    rq_activate_all_grippers(True)
    # end: URCap Program Node
  end
  $ 55 "zero_ftsensor()"
  zero_ftsensor()
  $ 56 "EXTT"
  $ 57 "Set GRP_3F_Enable=Off"
  set_standard_digital_out(4, False)
  $ 58 "Set BarcodeTrigger=Off"
  set_standard_digital_out(6, False)
  $ 59 "Set GRP_3F_Decap=Off"
  set_standard_digital_out(3, False)
  $ 60 "Set GRP_3F_Cap=Off"
  set_standard_digital_out(2, False)
  $ 61 "Set GRP_3F_Open=Off"
  set_standard_digital_out(5, False)
  $ 62 "PSE_T≔get_tool_free_pose(dir=[0,0,0.150], move_in_base_frame=True)"
  global PSE_T=get_tool_free_pose(dir=[0,0,0.150], move_in_base_frame=True)
  $ 63 "If is_reachable(Base_const, [PSE_T])"
  if (is_reachable(p[0.0,0.0,0.0,0.0,0.0,0.0], [PSE_T])):
    $ 64 "MoveL"
    $ 65 "PSE_T" "breakAfter"
    movel(PSE_T, a=1.2, v=0.15)
  end
  while (True):
    $ 66 "Robot Program"
    $ 67 "MAIN"
    $ 68 "command_manager(external_control='uGO', cond_suspend=(ITM_Manipulated and AMR_AtTarget and AMR_Charging and AMR_Battery<40), cond_unsuspend=(AMR_Battery≟60))"
    command_manager(external_control="uGO", cond_suspend=(ITM_Manipulated  and  AMR_AtTarget  and  AMR_Charging  and  AMR_Battery<40), cond_unsuspend=(AMR_Battery == 60))
    $ 69 "log_state(STATE_Info)"
    log_state(STATE_Info)
    $ 70 "Switch STATE"
    switch_1 = STATE
    $ 71 "Case 1"
    if (1 == switch_1):
      $ 72 "Stopping"
      $ 73 "STATE_Info≔'Stopping'"
      global STATE_Info="Stopping"
      $ 74 "end_freedrive_mode()"
      end_freedrive_mode()
      $ 75 "Set"
      set_tcp(p[0.0,0.0,0.161,3.1415,0.0,0.0])
      $ 76 "PSE_T≔get_tool_free_pose(dir=[0,0,0.150], move_in_base_frame=True)"
      global PSE_T=get_tool_free_pose(dir=[0,0,0.150], move_in_base_frame=True)
      $ 77 "If is_reachable(Base_const, [PSE_T])"
      if (is_reachable(p[0.0,0.0,0.0,0.0,0.0,0.0], [PSE_T])):
        $ 78 "MoveL"
        $ 79 "PSE_T" "breakAfter"
        movel(PSE_T, a=1.2, v=0.15)
      end
      $ 80 "do_transition(keep_rxry=OBJ_Picked, r=0)"
      do_transition(keep_rxry=OBJ_Picked, r=0)
      $ 89 "Call Sub_AMR_MiR_V3"
      Sub_AMR_MiR_V3()
      $ 90 "If stopping() and AMR_Done"
      if (stopping()  and  AMR_Done):
        $ 91 "STATE≔2"
        global STATE=2
        $ 92 "ugo_update_outputs()"
        ugo_update_outputs()
      end
    elif (2 == switch_1):
      $ 93 "Case 2"
      $ 94 "Stopped"
      $ 95 "STATE_Info≔'Stopped'"
      global STATE_Info="Stopped"
      $ 96 "Call Sub_AMR_MiR_V3"
      Sub_AMR_MiR_V3()
      $ 97 "If CMD_Reset"
      if (CMD_Reset):
        $ 98 "STATE≔3"
        global STATE=3
        $ 99 "ugo_update_outputs()"
        ugo_update_outputs()
      end
    elif (3 == switch_1):
      $ 100 "Case 3"
      $ 101 " Resetting"
      $ 102 "STATE_Info≔'Resetting'"
      global STATE_Info="Resetting"
      $ 103 "uML"
      $ 104 "reset_error()"
      reset_error()
      $ 105 "reset_warning()"
      reset_warning()
      $ 106 "PROCESS_Step≔0"
      global PROCESS_Step=0
      $ 107 "PROCESS_Info≔''"
      global PROCESS_Info=""
      $ 108 "ARM_Referenced≔ False "
      global ARM_Referenced=  False
      $ 109 "WRK_Done≔ False "
      global WRK_Done=  False
      $ 110 "ITM_Prepared≔ False "
      global ITM_Prepared=  False
      $ 111 "ITM_Manipulated≔ False "
      global ITM_Manipulated=  False
      $ 112 "STP≔0"
      global STP=0
      $ 113 "Action≔0"
      global Action=0
      $ 114 "Action_Info≔''"
      global Action_Info=""
      $ 115 "ITM_ID≔0"
      global ITM_ID=0
      $ 116 "JIG≔0"
      global JIG=0
      $ 117 "JIG_Slot≔0"
      global JIG_Slot=0
      $ 118 "Task_info≔''"
      global Task_info=""
      $ 119 "Set"
      set_tcp(p[0.0,0.0,0.161,3.1415,0.0,0.0])
      $ 120 "App"
      $ 121 "'ADD APPLICATION SPECIFIC COMMANDS'"
      # 'ADD APPLICATION SPECIFIC COMMANDS'
      $ 122 "OBJ_Type≔0"
      global OBJ_Type=0
      $ 123 "OBJ_Nbr≔0"
      global OBJ_Nbr=0
      $ 124 "If CNT_Rack_Output≥50"
      if (CNT_Rack_Output >= 50):
        $ 125 "CNT_Rack_Output≔0"
        global CNT_Rack_Output=0
      end
      $ 126 "TASK≔struct(ID=0, NAVI=struct(target=0, footprint=0, protectiveOff=0, dock=0), WORK=struct(ITM_ID_Src=0, JIG_ID_Src=0, OBJ_Nbr_Src=0, ACT_Src=0, ITM_ID_Tgt=0, JIG_ID_Tgt=0, OBJ_Nbr_Tgt=0, ACT_Tgt=0, OBJ_Type=0))"
      global TASK=struct(ID=0, NAVI=struct(target=0, footprint=0, protectiveOff=0, dock=0), WORK=struct(ITM_ID_Src=0, JIG_ID_Src=0, OBJ_Nbr_Src=0, ACT_Src=0, ITM_ID_Tgt=0, JIG_ID_Tgt=0, OBJ_Nbr_Tgt=0, ACT_Tgt=0, OBJ_Type=0))
      $ 127 "Call Sub_AMR_MiR_V3"
      Sub_AMR_MiR_V3()
      $ 128 "If resetting() and AMR_Done"
      if (resetting()  and  AMR_Done):
        $ 129 "STATE≔4"
        global STATE=4
        $ 130 "ugo_update_outputs()"
        ugo_update_outputs()
      end
    elif (4 == switch_1):
      $ 131 "Case 4"
      $ 132 "Idle"
      $ 133 "STATE_Info≔'Idle'"
      global STATE_Info="Idle"
      $ 134 "If CMD_Start"
      if (CMD_Start):
        $ 135 "STATE≔5"
        global STATE=5
        $ 136 "ugo_update_outputs()"
        ugo_update_outputs()
      end
    elif (5 == switch_1):
      $ 137 "Case 5"
      $ 138 "Starting"
      $ 139 "STATE_Info≔'Starting'"
      global STATE_Info="Starting"
      $ 140 "'ADD COMMANDS WHAT TO START WITH'"
      # 'ADD COMMANDS WHAT TO START WITH'
      $ 141 "Call Sub_AMR_MiR_V3"
      Sub_AMR_MiR_V3()
      $ 142 "get ugo data"
      $ 143 "Assign Tasks"
      $ 144 "TASK.ID = ugo_get_task()"
      TASK.ID = ugo_get_task()
      $ 145 "If TASK.ID≟1"
      if (TASK.ID == 1):
        $ 146 "Task_info≔'Charge'"
        global Task_info="Charge"
        $ 147 "Parameters"
        $ 148 "AMR_PosTarget≔1"
        global AMR_PosTarget=1
      else:
        $ 149 "ElseIf TASK.ID≟9"
        if (TASK.ID == 9):
          $ 150 "'Pick Sarstedt Rack from Variable source'"
          # 'Pick Sarstedt Rack from Variable source'
          $ 151 "Task_info≔'Navigate to Target'"
          global Task_info="Navigate to Target"
          $ 152 "Parameters"
          $ 153 "AMR_PosTarget≔UGO.read_input('00','ITM_ID')"
          global AMR_PosTarget=UGO.read_input("00","ITM_ID")
        else:
          $ 154 "ElseIf TASK.ID≟10"
          if (TASK.ID == 10):
            $ 155 "'Pick Sarstedt Rack from Variable source'"
            # 'Pick Sarstedt Rack from Variable source'
            $ 156 "Task_info≔'Pick Rack'"
            global Task_info="Pick Rack"
            $ 157 "AMR_PosTarget≔2"
            global AMR_PosTarget=2
            $ 158 "Parameters"
            $ 159 "ITM_ID≔UGO.read_input('00','ITM_ID')"
            global ITM_ID=UGO.read_input("00","ITM_ID")
            $ 160 "JIG≔UGO.read_input('00','JIG_ID')"
            global JIG=UGO.read_input("00","JIG_ID")
            $ 161 "OBJ_Type≔3"
            global OBJ_Type=3
          else:
            $ 162 "ElseIf TASK.ID≟11"
            if (TASK.ID == 11):
              $ 163 "'Place Sarstedt Rack on Variable target'"
              # 'Place Sarstedt Rack on Variable target'
              $ 164 "Task_info≔'Place Rack'"
              global Task_info="Place Rack"
              $ 165 "AMR_PosTarget≔2"
              global AMR_PosTarget=2
              $ 166 "Parameters"
              $ 167 "ITM_ID≔UGO.read_input('00','ITM_ID')"
              global ITM_ID=UGO.read_input("00","ITM_ID")
              $ 168 "JIG≔UGO.read_input('00','JIG_ID')"
              global JIG=UGO.read_input("00","JIG_ID")
              $ 169 "OBJ_Type≔3"
              global OBJ_Type=3
            else:
              $ 171 "ElseIf TASK.ID≟12"
              if (TASK.ID == 12):
                $ 172 "Task_info≔'Decapping'"
                global Task_info="Decapping"
                $ 173 "Parameters"
                $ 174 "ITM_ID≔1"
                global ITM_ID=1
                $ 175 "AMR_PosTarget≔AMR_PosActual"
                global AMR_PosTarget=AMR_PosActual
                $ 176 "PRC_TubCounter≔0"
                global PRC_TubCounter=0
              else:
                $ 177 "ElseIf TASK.ID≟13"
                if (TASK.ID == 13):
                  $ 178 "Task_info≔'Empty racks'"
                  global Task_info="Empty racks"
                  $ 179 "Parameters"
                  $ 180 "ITM_ID≔1"
                  global ITM_ID=1
                  $ 181 "AMR_PosTarget≔AMR_PosActual"
                  global AMR_PosTarget=AMR_PosActual
                else:
                  $ 182 "ElseIf TASK.ID≟16"
                  if (TASK.ID == 16):
                    $ 183 "Task_info≔'Decap + Barcode'"
                    global Task_info="Decap + Barcode"
                    $ 184 "Parameters"
                    $ 186 "OBJs_String≔UGO.read_input('00','ObjPos')"
                    global OBJs_String=UGO.read_input("00","ObjPos")
                    $ 187 "OBJs_List≔make_list(length = elements_in_string(OBJs_String), initial_value = -1, capacity = 50)"
                    global OBJs_List=make_list(length = elements_in_string(OBJs_String), initial_value = -1, capacity = 50)
                    $ 188 "OBJs_List≔string_to_list(OBJs_String)"
                    global OBJs_List=string_to_list(OBJs_String)
                    $ 189 "ITM_ID≔1"
                    global ITM_ID=1
                    $ 190 "OBJ_Type≔2"
                    global OBJ_Type=2
                    $ 191 "JIG≔7"
                    global JIG=7
                    $ 192 "AMR_PosTarget≔AMR_PosActual"
                    global AMR_PosTarget=AMR_PosActual
                  else:
                    $ 193 "ElseIf TASK.ID≟99"
                    if (TASK.ID == 99):
                      $ 194 "Task_info≔'Decapping and barcode alignment'"
                      global Task_info="Decapping and barcode alignment"
                      $ 195 "Parameters"
                      $ 196 "PRC_TubNumber≔UGO.read_input('00','TubesNb')"
                      global PRC_TubNumber=UGO.read_input("00","TubesNb")
                      $ 197 "PRC_TubCounter≔0"
                      global PRC_TubCounter=0
                      $ 198 "ITM_ID≔1"
                      global ITM_ID=1
                      $ 199 "AMR_PosTarget≔AMR_PosActual"
                      global AMR_PosTarget=AMR_PosActual
                    else:
                      $ 234 "Else" "noBreak"
                      $ 235 "set_error(ERROR_WRONG_ORDER)"
                      set_error(ERROR_WRONG_ORDER)
                    end
                  end
                end
              end
            end
          end
        end
      end
      $ 236 "test ugo"
      $ 237 "Wait: 0.2"
      sleep(0.2)
      $ 238 "ugo_update_outputs()"
      ugo_update_outputs()
      $ 239 "If starting() and AMR_Done"
      if (starting()  and  AMR_Done):
        $ 240 "log_message(Task_info, 'New Task: ')"
        log_message(Task_info, "New Task: ")
        $ 241 "log_message(to_str(TASK.ID), 'Task_ID: ')"
        log_message(to_str(TASK.ID), "Task_ID: ")
        $ 242 "do_transition(keep_rxry=OBJ_Picked)"
        do_transition(keep_rxry=OBJ_Picked)
        $ 243 "STATE≔6"
        global STATE=6
        $ 244 "ugo_update_outputs()"
        ugo_update_outputs()
      end
    elif (6 == switch_1):
      $ 245 "Case 6"
      $ 246 "Execute"
      $ 247 "STATE_Info≔'Execute'"
      global STATE_Info="Execute"
      $ 248 "If  not CMD_Hold and not CMD_Suspend"
      global thread_flag_248=0
      thread Thread_if_248():
        $ 249 "Switch PROCESS_Step"
        switch_2 = PROCESS_Step
        $ 250 "Case 0"
        if (0 == switch_2):
          $ 251 "PROCESS_Info≔'process control'"
          global PROCESS_Info="process control"
          $ 252 "log_process(PROCESS_Info)"
          log_process(PROCESS_Info)
          $ 253 "process control"
          $ 254 "If  not AMR_AtTarget"
          if (  not  AMR_AtTarget):
            $ 255 "PROCESS_Step≔1"
            global PROCESS_Step=1
          else:
            $ 256 "ElseIf (( not ITM_Prepared and  not WRK_Done) or (ITM_Prepared and WRK_Done))"
            if (((  not  ITM_Prepared  and    not  WRK_Done)  or  (ITM_Prepared  and  WRK_Done))):
              $ 257 "PROCESS_Step≔2"
              global PROCESS_Step=2
            else:
              $ 258 "ElseIf  not WRK_Done"
              if (  not  WRK_Done):
                $ 259 "PROCESS_Step≔3"
                global PROCESS_Step=3
              else:
                $ 260 "Else" "noBreak"
                $ 261 "task finished"
                $ 262 "PROCESS_Info≔''"
                global PROCESS_Info=""
                $ 263 "STATE≔7"
                global STATE=7
                $ 264 "ugo_update_outputs()"
                ugo_update_outputs()
              end
            end
          end
        elif (1 == switch_2):
          $ 265 "Case 1"
          $ 266 "navigate"
          $ 267 "'MOVING THE uML'"
          # 'MOVING THE uML'
          $ 268 "PROCESS_Info≔'move to target'"
          global PROCESS_Info="move to target"
          $ 269 "log_process(PROCESS_Info)"
          log_process(PROCESS_Info)
          $ 270 "If TASK.ID≟1"
          if (TASK.ID == 1):
            $ 271 "Action≔51"
            global Action=51
          else:
            $ 272 "Else" "noBreak"
            $ 273 "Action≔52"
            global Action=52
          end
          $ 274 "Call Sub_AMR_MiR_V3"
          Sub_AMR_MiR_V3()
          $ 275 "If AMR_Done"
          if (AMR_Done):
            $ 276 "PROCESS_Step≔0"
            global PROCESS_Step=0
          end
        elif (2 == switch_2):
          $ 277 "Case 2"
          $ 278 "prepare"
          $ 279 "'THINGS THAT HAVE TO BE DONE ONCE IN A SEQUENCE,WORKFLOW'"
          # 'THINGS THAT HAVE TO BE DONE ONCE IN A SEQUENCE,WORKFLOW'
          $ 280 "PROCESS_Info≔'prepare for work'"
          global PROCESS_Info="prepare for work"
          $ 281 "log_process(PROCESS_Info)"
          log_process(PROCESS_Info)
          $ 282 "If TASK.WORK.ITM_ID_Src>1"
          if (TASK.WORK.ITM_ID_Src>1):
            $ 283 "ITM_ID≔TASK.WORK.ITM_ID_Src"
            global ITM_ID=TASK.WORK.ITM_ID_Src
          else:
            $ 284 "ElseIf TASK.WORK.ITM_ID_Tgt>1"
            if (TASK.WORK.ITM_ID_Tgt>1):
              $ 285 "ITM_ID≔TASK.WORK.ITM_ID_Tgt"
              global ITM_ID=TASK.WORK.ITM_ID_Tgt
            end
          end
          $ 286 "If  not ARM_Referenced and (ITM_ID≠0)"
          if (  not  ARM_Referenced  and  (ITM_ID != 0)):
            $ 287 "STP≔1"
            global STP=1
          else:
            $ 288 "ElseIf ARM_Referenced or (ITM_ID≟0)"
            if (ARM_Referenced  or  (ITM_ID == 0)):
              $ 289 "STP≔2"
              global STP=2
            end
          end
          $ 290 "Switch STP"
          switch_3 = STP
          $ 291 "Case 1"
          if (1 == switch_3):
            $ 292 "reference"
            $ 293 "STP_Info≔'reference at target position'"
            global STP_Info="reference at target position"
            $ 294 "log_step(STP_Info)"
            log_step(STP_Info)
            $ 295 "If ITM_ID≟1"
            if (ITM_ID == 1):
              $ 296 "CAM_Done≔ True "
              global CAM_Done=  True
            else:
              $ 297 "Else" "noBreak"
              $ 298 "Action≔131"
              global Action=131
              $ 299 "Call Sub_Vision_V18"
              Sub_Vision_V18()
            end
            $ 301 "If CAM_Done and  not ERROR.FLAG"
            if (CAM_Done  and    not  ERROR.FLAG):
              $ 302 "log_step('ARM referenced')"
              log_step("ARM referenced")
              $ 303 "ARM_Referenced≔ True "
              global ARM_Referenced=  True
            end
          elif (2 == switch_3):
            $ 304 "Case 2"
            $ 305 "manipulate"
            $ 306 "STP_Info≔'manipulate item'"
            global STP_Info="manipulate item"
            $ 307 "log_step(STP_Info)"
            log_step(STP_Info)
            $ 308 "'In case pressing button is needed'"
            # 'In case pressing button is needed'
            $ 309 "If found_in_list(ITM_ID, ITM_ID_List)"
            if (found_in_list(ITM_ID, ITM_ID_List)):
              $ 310 "Switch ITM_ID"
              switch_4 = ITM_ID
              $ 311 "Case 0"
              if (0 == switch_4):
                $ 312 "ITM_Manipulated≔ not ITM_Manipulated"
                global ITM_Manipulated=  not  ITM_Manipulated
              elif (1 == switch_4):
                $ 313 "Case 1"
                $ 314 "ITM_Manipulated≔ not ITM_Manipulated"
                global ITM_Manipulated=  not  ITM_Manipulated
              elif (2 == switch_4):
                $ 315 "Case 2"
              else:
                $ 325 "Default Case"
                $ 326 "ITM_Manipulated≔ not ITM_Manipulated"
                global ITM_Manipulated=  not  ITM_Manipulated
              end
            end
          end
          $ 327 "ITM_Prepared≔(ITM_Manipulated or  not found_in_list(ITM_ID, ITM_ID_List)) and (ARM_Referenced or ITM_ID≟0) and  not WRK_Done"
          global ITM_Prepared=(ITM_Manipulated  or    not  found_in_list(ITM_ID, ITM_ID_List))  and  (ARM_Referenced  or  ITM_ID == 0)  and    not  WRK_Done
          $ 328 "STP≔0"
          global STP=0
          $ 329 "STP_Info≔''"
          global STP_Info=""
          $ 330 "PROCESS_Step≔0"
          global PROCESS_Step=0
        elif (3 == switch_2):
          $ 331 "Case 3"
          $ 332 "work"
          $ 333 "'ADD EVERY MACHINE, OBJECT, STATION TO WORK ON'"
          # 'ADD EVERY MACHINE, OBJECT, STATION TO WORK ON'
          $ 334 "Switch ITM_ID"
          switch_3 = ITM_ID
          $ 335 "Case 1"
          if (1 == switch_3):
            $ 336 "uLM"
            $ 337 "If TASK.ID≟12"
            if (TASK.ID == 12):
              $ 338 "fill racks"
              $ 339 "Action≔151"
              global Action=151
              $ 340 "Call Sub_Vision_V18"
              Sub_Vision_V18()
              $ 341 "If  not ERROR.FLAG"
              if (  not  ERROR.FLAG):
                $ 342 "Actions for the task"
                $ 343 "Action≔1"
                global Action=1
                $ 344 "JIG≔2"
                global JIG=2
                $ 345 "JIG_Slot≔CAM_Result[0]"
                global JIG_Slot=CAM_Result[0]
                $ 346 "OBJ_Nbr≔CAM_Result[0]"
                global OBJ_Nbr=CAM_Result[0]
                $ 347 "OBJ_Type≔2"
                global OBJ_Type=2
                $ 348 "Call Sub_Action_V4"
                Sub_Action_V4()
                $ 349 "If OBJ_Picked"
                if (OBJ_Picked):
                  $ 350 "CAM_Result.remove(0)"
                  CAM_Result.remove(0)
                  $ 351 "PRC_TubCounter≔PRC_TubCounter+1"
                  global PRC_TubCounter=PRC_TubCounter+1
                  $ 352 "If PRC_TubCounter%4≟0"
                  if (PRC_TubCounter%4 == 0):
                    $ 353 "JIG_Slot≔4"
                    global JIG_Slot=4
                  else:
                    $ 354 "Else" "noBreak"
                    $ 355 "JIG_Slot≔PRC_TubCounter%4"
                    global JIG_Slot=PRC_TubCounter%4
                  end
                  $ 356 "OBJ_Nbr≔ceil(PRC_TubCounter/4)"
                  global OBJ_Nbr=ceil(PRC_TubCounter/4)
                  $ 357 "Action≔2"
                  global Action=2
                  $ 358 "JIG≔4"
                  global JIG=4
                  $ 359 "Call Sub_Action_V4"
                  Sub_Action_V4()
                  $ 360 "Action≔151"
                  global Action=151
                  $ 361 "Call Sub_Vision_V18"
                  Sub_Vision_V18()
                end
              end
              $ 362 "If (CAM_Captures≥CAM_PRM_Retries) or (PRC_TubCounter≥32)"
              if ((CAM_Captures >= CAM_PRM_Retries)  or  (PRC_TubCounter >= 32)):
                $ 363 "PROCESS_Step≔0"
                global PROCESS_Step=0
                $ 364 "WRK_Done≔ True "
                global WRK_Done=  True
              end
            else:
              $ 365 "ElseIf TASK.ID≟10"
              if (TASK.ID == 10):
                $ 366 "Pick Rack"
                $ 367 "Action≔131"
                global Action=131
                $ 368 "Call Sub_Vision_V18"
                Sub_Vision_V18()
                $ 369 "Action≔1"
                global Action=1
                $ 370 "Call Sub_Action_V4"
                Sub_Action_V4()
                $ 371 "PROCESS_Step≔0"
                global PROCESS_Step=0
                $ 372 "WRK_Done≔ True "
                global WRK_Done=  True
              else:
                $ 373 "ElseIf TASK.ID≟11"
                if (TASK.ID == 11):
                  $ 374 "Place Rack"
                  $ 375 "Action≔2"
                  global Action=2
                  $ 376 "Call Sub_Action_V4"
                  Sub_Action_V4()
                  $ 377 "PROCESS_Step≔0"
                  global PROCESS_Step=0
                  $ 378 "WRK_Done≔ True "
                  global WRK_Done=  True
                else:
                  $ 379 "ElseIf TASK.ID≟13"
                  if (TASK.ID == 13):
                    $ 380 "empty racks"
                    $ 381 "pick"
                    $ 382 "Action≔1"
                    global Action=1
                    $ 383 "JIG≔4"
                    global JIG=4
                    $ 384 "If PRC_TubCounter%4≟0"
                    if (PRC_TubCounter%4 == 0):
                      $ 385 "JIG_Slot≔4"
                      global JIG_Slot=4
                    else:
                      $ 386 "Else" "noBreak"
                      $ 387 "JIG_Slot≔PRC_TubCounter%4"
                      global JIG_Slot=PRC_TubCounter%4
                    end
                    $ 388 "OBJ_Nbr≔ceil(PRC_TubCounter/4)"
                    global OBJ_Nbr=ceil(PRC_TubCounter/4)
                    $ 389 "OBJ_Type≔2"
                    global OBJ_Type=2
                    $ 390 "Call Sub_Action_V4"
                    Sub_Action_V4()
                    $ 391 "If OBJ_Picked"
                    if (OBJ_Picked):
                      $ 392 "Action≔2"
                      global Action=2
                      $ 393 "JIG≔3"
                      global JIG=3
                      $ 394 "JIG_Slot≔1"
                      global JIG_Slot=1
                      $ 395 "CNT_Rack_Output≔CNT_Rack_Output + 1"
                      global CNT_Rack_Output=CNT_Rack_Output + 1
                      $ 396 "OBJ_Nbr≔CNT_Rack_Output"
                      global OBJ_Nbr=CNT_Rack_Output
                      $ 397 "Call Sub_Action_V4"
                      Sub_Action_V4()
                      $ 398 "If  not ERROR.FLAG"
                      if (  not  ERROR.FLAG):
                        $ 399 "PRC_TubCounter≔PRC_TubCounter - 1"
                        global PRC_TubCounter=PRC_TubCounter - 1
                      end
                    end
                    $ 400 "If CNT_Rack_Output≥50 or PRC_TubCounter≤0"
                    if (CNT_Rack_Output >= 50  or  PRC_TubCounter <= 0):
                      $ 401 "PROCESS_Step≔0"
                      global PROCESS_Step=0
                      $ 402 "WRK_Done≔ True "
                      global WRK_Done=  True
                    end
                  else:
                    $ 403 "ElseIf TASK.ID≟16"
                    if (TASK.ID == 16):
                      $ 404 "CAM_Result≔OBJs_List"
                      global CAM_Result=OBJs_List
                      $ 405 "PRC_CntDetect≔0"
                      global PRC_CntDetect=0
                      $ 406 "Loop PRC_CntDetect<CAM_Result.length()"
                      while (PRC_CntDetect<CAM_Result.length()):
                        $ 407 "Action≔1"
                        global Action=1
                        $ 408 "ITM_ID≔1"
                        global ITM_ID=1
                        $ 409 "JIG≔2"
                        global JIG=2
                        $ 410 "OBJ_Type≔2"
                        global OBJ_Type=2
                        $ 411 "JIG_Slot≔CAM_Result[PRC_CntDetect]"
                        global JIG_Slot=CAM_Result[PRC_CntDetect]
                        $ 412 "OBJ_Nbr≔CAM_Result[PRC_CntDetect]"
                        global OBJ_Nbr=CAM_Result[PRC_CntDetect]
                        $ 413 "Call Sub_Action_V4"
                        Sub_Action_V4()
                        $ 414 "JIG≔1"
                        global JIG=1
                        $ 415 "Action≔11"
                        global Action=11
                        $ 416 "Call Sub_Action_V4"
                        Sub_Action_V4()
                        $ 417 "Action≔12"
                        global Action=12
                        $ 418 "Call Sub_Action_V4"
                        Sub_Action_V4()
                        $ 419 "Action≔6"
                        global Action=6
                        $ 420 "JIG≔6"
                        global JIG=6
                        $ 421 "Call Sub_Action_V4"
                        Sub_Action_V4()
                        $ 422 "Action≔13"
                        global Action=13
                        $ 423 "Call Sub_Action_V4"
                        Sub_Action_V4()
                        $ 424 "Action≔1"
                        global Action=1
                        $ 425 "JIG≔1"
                        global JIG=1
                        $ 426 "Call Sub_Action_V4"
                        Sub_Action_V4()
                        $ 427 "If OBJ_Brc_OK"
                        if (OBJ_Brc_OK):
                          $ 428 "JIG≔2"
                          global JIG=2
                          $ 429 "Action≔2"
                          global Action=2
                          $ 430 "OBJ_Nbr≔CAM_Result[PRC_CntDetect]"
                          global OBJ_Nbr=CAM_Result[PRC_CntDetect]
                          $ 431 "JIG_Slot≔CAM_Result[PRC_CntDetect]"
                          global JIG_Slot=CAM_Result[PRC_CntDetect]
                          $ 432 "OBJ_Type≔2"
                          global OBJ_Type=2
                          $ 433 "Call Sub_Action_V4"
                          Sub_Action_V4()
                        else:
                          $ 434 "Else" "noBreak"
                          $ 435 "Action≔2"
                          global Action=2
                          $ 436 "JIG≔8"
                          global JIG=8
                          $ 437 "Call Sub_Action_V4"
                          Sub_Action_V4()
                        end
                        $ 438 "PRC_CntDetect≔PRC_CntDetect+1"
                        global PRC_CntDetect=PRC_CntDetect+1
                      end
                      $ 439 "PROCESS_Step≔0"
                      global PROCESS_Step=0
                      $ 440 "WRK_Done≔ True "
                      global WRK_Done=  True
                    end
                  end
                end
              end
            end
          elif (2 == switch_3):
            $ 441 "Case 2"
          elif (5 == switch_3):
            $ 483 "Case 5"
            $ 484 "SarstedtTable"
            $ 485 "Action≔131"
            global Action=131
            $ 486 "Call Sub_Vision_V18"
            Sub_Vision_V18()
            $ 487 "Action≔1"
            global Action=1
            $ 488 "Call Sub_Action_V4"
            Sub_Action_V4()
            $ 489 "PROCESS_Step≔0"
            global PROCESS_Step=0
            $ 490 "WRK_Done≔ True "
            global WRK_Done=  True
          elif (20 == switch_3):
            $ 491 "Case 20"
          else:
            $ 553 "Default Case"
            $ 554 "WRK_Done≔ True "
            global WRK_Done=  True
            $ 555 "PROCESS_Step≔0"
            global PROCESS_Step=0
          end
        end
        thread_flag_248 = 1
      end
      if (  not  CMD_Hold and not CMD_Suspend):
        global thread_handler_248=run Thread_if_248()
        while (thread_flag_248 == 0):
          if not(  not  CMD_Hold and not CMD_Suspend):
            kill thread_handler_248
            thread_flag_248 = 2
          else:
            sync()
          end
        end
      else:
        thread_flag_248 = 2
      end
      $ 556 "If CMD_Hold"
      if (CMD_Hold):
        $ 557 "STATE≔9"
        global STATE=9
        $ 558 "ugo_update_outputs()"
        ugo_update_outputs()
      else:
        $ 559 "ElseIf CMD_Suspend"
        if (CMD_Suspend):
          $ 560 "STATE≔12"
          global STATE=12
          $ 561 "ugo_update_outputs()"
          ugo_update_outputs()
        end
      end
    elif (7 == switch_1):
      $ 562 "Case 7"
      $ 563 "Completing"
      $ 564 "STATE_Info≔'Completing'"
      global STATE_Info="Completing"
      $ 565 "'ADD COMMANDS FOR COMPLETING THE PROCESS'"
      # 'ADD COMMANDS FOR COMPLETING THE PROCESS'
      $ 566 "do_transition(keep_rxry=OBJ_Picked)"
      do_transition(keep_rxry=OBJ_Picked)
      $ 567 "Call Sub_AMR_MiR_V3"
      Sub_AMR_MiR_V3()
      $ 568 "If completing() and AMR_Done"
      if (completing()  and  AMR_Done):
        $ 569 "STATE≔8"
        global STATE=8
        $ 570 "ugo_update_outputs()"
        ugo_update_outputs()
      end
    elif (8 == switch_1):
      $ 571 "Case 8"
      $ 572 "Complete"
      $ 573 "STATE_Info≔'Complete'"
      global STATE_Info="Complete"
      $ 574 "If CMD_Reset"
      if (CMD_Reset):
        $ 575 "STATE≔3"
        global STATE=3
        $ 576 "ugo_update_outputs()"
        ugo_update_outputs()
      end
    elif (9 == switch_1):
      $ 577 "Case 9"
      $ 578 "Holding"
      $ 579 "STATE_Info≔'Holding'"
      global STATE_Info="Holding"
      $ 580 "stopl(0.5)"
      stopl(0.5)
      $ 581 "Call Sub_AMR_MiR_V3"
      Sub_AMR_MiR_V3()
      $ 582 "If holding() and AMR_Done"
      if (holding()  and  AMR_Done):
        $ 583 "STATE≔10"
        global STATE=10
        $ 584 "ugo_update_outputs()"
        ugo_update_outputs()
      end
    elif (10 == switch_1):
      $ 585 "Case 10"
      $ 586 "Held"
      $ 587 "STATE_Info≔'Held'"
      global STATE_Info="Held"
      $ 588 "If CMD_Unhold"
      if (CMD_Unhold):
        $ 589 "end_freedrive_mode()"
        end_freedrive_mode()
        $ 590 "STATE≔11"
        global STATE=11
        $ 591 "ugo_update_outputs()"
        ugo_update_outputs()
      else:
        $ 592 "ElseIf FNC_Freedrive"
        if (FNC_Freedrive):
          $ 593 "freedrive_mode()"
          freedrive_mode()
        else:
          $ 594 "Else" "noBreak"
          $ 595 "end_freedrive_mode()"
          end_freedrive_mode()
        end
      end
    elif (11 == switch_1):
      $ 596 "Case 11"
      $ 597 "Unholding"
      $ 598 "STATE_Info≔'Unholding'"
      global STATE_Info="Unholding"
      $ 599 "Clearing"
      $ 600 "Switch ERROR.ID"
      switch_2 = ERROR.ID
      $ 601 "Case 1002"
      if (1002 == switch_2):
        $ 602 "AMR_AtTarget≔ False "
        global AMR_AtTarget=  False
        $ 603 "ARM_Referenced≔ False "
        global ARM_Referenced=  False
        $ 604 "ITM_Prepared≔ False "
        global ITM_Prepared=  False
        $ 605 "PROCESS_Step≔1"
        global PROCESS_Step=1
      elif (2007 == switch_2):
        $ 606 "Case 2007"
        $ 607 "PROCESS_Step≔1"
        global PROCESS_Step=1
      end
      $ 608 "reset_error()"
      reset_error()
      $ 609 "reset_warning()"
      reset_warning()
      $ 610 "OBJ_Picked≔gripper_has_object()"
      global OBJ_Picked=gripper_has_object()
      $ 611 "Call Sub_AMR_MiR_V3"
      Sub_AMR_MiR_V3()
      $ 612 "If unholding() and AMR_Done"
      if (unholding()  and  AMR_Done):
        $ 613 "STATE≔6"
        global STATE=6
        $ 614 "ugo_update_outputs()"
        ugo_update_outputs()
      end
    elif (12 == switch_1):
      $ 615 "Case 12"
      $ 616 "Suspending"
      $ 617 "STATE_Info≔'Suspending'"
      global STATE_Info="Suspending"
      $ 618 "PROCESS_Info≔str_cat(PROCESS_Info, ' suspended')"
      global PROCESS_Info=str_cat(PROCESS_Info, " suspended")
      $ 619 "If suspending()"
      if (suspending()):
        $ 620 "STATE≔13"
        global STATE=13
        $ 621 "ugo_update_outputs()"
        ugo_update_outputs()
      end
    elif (13 == switch_1):
      $ 622 "Case 13"
      $ 623 "Suspended"
      $ 624 "STATE_Info≔'Suspended'"
      global STATE_Info="Suspended"
      $ 625 "Call Sub_AMR_MiR_V3"
      Sub_AMR_MiR_V3()
      $ 626 "If CMD_Unsuspend"
      if (CMD_Unsuspend):
        $ 627 "STATE≔14"
        global STATE=14
        $ 628 "ugo_update_outputs()"
        ugo_update_outputs()
      end
    elif (14 == switch_1):
      $ 629 "Case 14"
      $ 630 "Unsuspending"
      $ 631 "STATE_Info≔'Unsuspending'"
      global STATE_Info="Unsuspending"
      $ 632 "PROCESS_Step≔0"
      global PROCESS_Step=0
      $ 633 "If unsuspending()"
      if (unsuspending()):
        $ 634 "STATE≔6"
        global STATE=6
        $ 635 "ugo_update_outputs()"
        ugo_update_outputs()
      end
    elif (15 == switch_1):
      $ 636 "Case 15"
      $ 637 "Aborting"
      $ 638 "STATE_Info≔'Aborting'"
      global STATE_Info="Aborting"
      $ 639 "If aborting()"
      if (aborting()):
        $ 640 "STATE≔16"
        global STATE=16
        $ 641 "ugo_update_outputs()"
        ugo_update_outputs()
      end
    elif (16 == switch_1):
      $ 642 "Case 16"
      $ 643 "Aborted"
      $ 644 "STATE_Info≔'Aborted'"
      global STATE_Info="Aborted"
      $ 645 "If CMD_Clear"
      if (CMD_Clear):
        $ 646 "STATE≔17"
        global STATE=17
        $ 647 "ugo_update_outputs()"
        ugo_update_outputs()
      end
    elif (17 == switch_1):
      $ 648 "Case 17"
      $ 649 "Clearing"
      $ 650 "STATE_Info≔'Clearing'"
      global STATE_Info="Clearing"
      $ 651 "Clearing"
      $ 652 "reset_warning()"
      reset_warning()
      $ 653 "reset_error()"
      reset_error()
      $ 654 "If clearing()"
      if (clearing()):
        $ 655 "STATE≔2"
        global STATE=2
        $ 656 "ugo_update_outputs()"
        ugo_update_outputs()
      end
    end
    $ 657 "log_state(STATE_Info)"
    log_state(STATE_Info)
    $ 658 "log_warning(WARNING.MSG)"
    log_warning(WARNING.MSG)
    $ 659 "log_error(ERROR.MSG)"
    log_error(ERROR.MSG)
    $ 660 "Times"
    $ 661 "Switch STATE"
    switch_1 = STATE
    $ 662 "Case 1"
    if (1 == switch_1):
      $ 663 "TM_St_Stopping≔get_time(STATE_Times[STATE-1])"
      global TM_St_Stopping=get_time(STATE_Times[STATE-1])
    elif (2 == switch_1):
      $ 664 "Case 2"
      $ 665 "TM_St_Stopped≔get_time(STATE_Times[STATE-1])"
      global TM_St_Stopped=get_time(STATE_Times[STATE-1])
    elif (3 == switch_1):
      $ 666 "Case 3"
      $ 667 "TM_St_Resetting≔get_time(STATE_Times[STATE-1])"
      global TM_St_Resetting=get_time(STATE_Times[STATE-1])
    elif (4 == switch_1):
      $ 668 "Case 4"
      $ 669 "TM_St_Idle≔get_time(STATE_Times[STATE-1])"
      global TM_St_Idle=get_time(STATE_Times[STATE-1])
    elif (5 == switch_1):
      $ 670 "Case 5"
      $ 671 "TM_St_Starting≔get_time(STATE_Times[STATE-1])"
      global TM_St_Starting=get_time(STATE_Times[STATE-1])
    elif (6 == switch_1):
      $ 672 "Case 6"
      $ 673 "TM_St_Execute≔get_time(STATE_Times[STATE-1])"
      global TM_St_Execute=get_time(STATE_Times[STATE-1])
    elif (7 == switch_1):
      $ 674 "Case 7"
      $ 675 "TM_St_Completin≔get_time(STATE_Times[STATE-1])"
      global TM_St_Completin=get_time(STATE_Times[STATE-1])
    elif (8 == switch_1):
      $ 676 "Case 8"
      $ 677 "TM_St_Complete≔get_time(STATE_Times[STATE-1])"
      global TM_St_Complete=get_time(STATE_Times[STATE-1])
    elif (9 == switch_1):
      $ 678 "Case 9"
      $ 679 "TM_St_Holding≔get_time(STATE_Times[STATE-1])"
      global TM_St_Holding=get_time(STATE_Times[STATE-1])
    elif (10 == switch_1):
      $ 680 "Case 10"
      $ 681 "TM_St_Held≔get_time(STATE_Times[STATE-1])"
      global TM_St_Held=get_time(STATE_Times[STATE-1])
    elif (11 == switch_1):
      $ 682 "Case 11"
      $ 683 "TM_St_Unholding≔get_time(STATE_Times[STATE-1])"
      global TM_St_Unholding=get_time(STATE_Times[STATE-1])
    elif (12 == switch_1):
      $ 684 "Case 12"
      $ 685 "TM_St_Suspendin≔get_time(STATE_Times[STATE-1])"
      global TM_St_Suspendin=get_time(STATE_Times[STATE-1])
    elif (13 == switch_1):
      $ 686 "Case 13"
      $ 687 "TM_St_Suspended≔get_time(STATE_Times[STATE-1])"
      global TM_St_Suspended=get_time(STATE_Times[STATE-1])
    elif (14 == switch_1):
      $ 688 "Case 14"
      $ 689 "TM_St_Unsuspend≔get_time(STATE_Times[STATE-1])"
      global TM_St_Unsuspend=get_time(STATE_Times[STATE-1])
    elif (15 == switch_1):
      $ 690 "Case 15"
      $ 691 "TM_St_Aborting≔get_time(STATE_Times[STATE-1])"
      global TM_St_Aborting=get_time(STATE_Times[STATE-1])
    elif (16 == switch_1):
      $ 692 "Case 16"
      $ 693 "TM_St_Aborted≔get_time(STATE_Times[STATE-1])"
      global TM_St_Aborted=get_time(STATE_Times[STATE-1])
    elif (17 == switch_1):
      $ 694 "Case 17"
      $ 695 "TM_St_Clearing≔get_time(STATE_Times[STATE-1])"
      global TM_St_Clearing=get_time(STATE_Times[STATE-1])
    end
    $ 697 "Wait: 0.1"
    sleep(0.1)
  end
end
